VAR_GLOBAL
	bInletOpen		AT %Q*	: BOOL;
	bConveyorRun	AT %Q*	: BOOL;
	nLevelRaw		AT %I*	: INT;
	bStartButton	AT %I*	: BOOL;
	stDrive			AT %I*	: ST_DriveIn;
	aLamps			AT %Q*	: ARRAY[1..3] OF BOOL;
	bSpareOut		AT %Q*	: BOOL;	// spare: not linked
END_VAR

(* stored: Version 1.1.0.1
   GVL GVL_IO: Id {8a3bfc93-eaf8-4cd9-8dc2-625b6ff9b2c4} *)
